// TIA Portal V17 export
// export: Created 2025-07-10T10:56:05.3982501Z, ExportSetting WithDefaults, DisplayName Totally Integrated Automation Portal, DisplayVersion V17, DisplayName TIA Portal Openness, DisplayVersion V17, DisplayName TIA Portal Version Control Interface, DisplayVersion V17, DisplayName SINAMICS Startdrive Advanced, DisplayVersion V17, DisplayName SINAMICS Startdrive G130, G150, S120, S150, SINAMICS MV, S210, DisplayVersion V17, DisplayName SINAMICS Startdrive G110M, G120, G120C, G120D, G120P, G115D, DisplayVersion V17, DisplayName STEP 7 Professional, DisplayVersion V17, DisplayName STEP 7 Safety, DisplayVersion V17, DisplayName WinCC Professional, DisplayVersion V17
FUNCTION_BLOCK "PR_GantryUnload_Seqv2 5_d22cba"   // FB1, LAD
VERSION : 0.1
// stored: AutoNumber true, IsIECCheckEnabled false, UDAEnableTagReadback false
   VAR_INPUT
      iAutoRunning : Bool;
      iCenteringSlideAtHome : Bool;
      iDistSenHighLimit : Int;
      iDistSenLowLimit : Int;
      iDistSensorIP : Int;
      iDryCycleWithoutPal : Bool;
      iGantryOutofZone : Bool;
      iGantryPickOver : Bool;
      iPCAckZero : Bool;
      iPCBypass : Bool;
      iPCDataReadOver : Bool;
      iPCDataWriteOver : Bool;
      iPalletPresent : Bool;
      iProcessStart : Bool;
      iReset_fault : Bool;
      iRetryPB : Bool;
      iScanErr : Bool;
      iScanOver : Bool;
      iScannerBypass : Bool;
      iSstMode : Bool;
      iSstPB : Bool;
   END_VAR
   VAR_OUTPUT
      qCenteringSlideAdvance : Bool;
      qCenteringSlideRetract : Bool;
      qCheckDistance : Bool;
      qGantryOkToUnload : Bool;
      qMsg : Array[0..2] of Bool;
      qPCReadCmd : Bool;
      qPCUploadCmd : Bool;
      qProcessOver : Bool;
      qScanCmd : Bool;
   END_VAR
   VAR DB_SPECIFIC
      StateNo : Int;
      s44_WaitResetRelease : Bool;
      s44_WaitResetRelease_T1 : Bool;
      s45_WaitGantryOutZone : Bool;
      s45_WaitGantryOutZone_T1 : Bool;
      s46_ChkStationHome : Bool;
      s46_ChkStationHome_T1 : Bool;
      s46_ChkStationHome_T2 : Bool;
      s47_WaitProcStartPZR : Bool;
      s47_WaitProcStartPZR_T1 : Bool;
      s48_ChkRecovery : Bool;
      s48_ChkRecovery_T1 : Bool;
      s48_ChkRecovery_T2 : Bool;
      s48_ChkRecovery_T3 : Bool;
      s49_WaitCentSlideAdv : Bool;
      s49_WaitCentSlideAdv_T1 : Bool;
      s50_WaitDistSensorFB : Bool;
      s50_WaitDistSensorFB_T1 : Bool;
      s51_WaitCentSlideRet : Bool;
      s51_WaitCentSlideRet_T1 : Bool;
      s52_WaitScanOver : Bool;
      s52_WaitScanOver_T1 : Bool;
      s52_WaitScanOver_T2 : Bool;
      s53_ChkMeasDistPCDat : Bool;
      s53_ChkMeasDistPCDat_T1 : Bool;
      s53_ChkMeasDistPCDat_T2 : Bool;
      s54_WaitGantryUnload : Bool;
      s54_WaitGantryUnload_T1 : Bool;
      s55_WaitGantryUnldOvr : Bool;
      s55_WaitGantryUnldOvr_T1 : Bool;
      s56_WaitGantryOutZone : Bool;
      s56_WaitGantryOutZone_T1 : Bool;
      s57_ChkReelAbsentCnv : Bool;
      s57_ChkReelAbsentCnv_T1 : Bool;
      s58_WaitProcStartLow : Bool;
      s58_WaitProcStartLow_T1 : Bool;
      s61_ChkMeasDiamTol : Bool;
      s61_ChkMeasDiamTol_T1 : Bool;
      s61_ChkMeasDiamTol_T2 : Bool;
      s62_WaitPCAckZero : Bool;
      s62_WaitPCAckZero_T1 : Bool;
      s63_WaitDataWritePC : Bool;
      s63_WaitDataWritePC_T1 : Bool;
      s64_WaitOperatorIntv : Bool;
      s64_WaitOperatorIntv_T1 : Bool;
      s65_ChkScanRetryOver : Bool;
      s65_ChkScanRetryOver_T1 : Bool;
      s65_ChkScanRetryOver_T2 : Bool;
      s66_WaitOperatorDecn : Bool;
      s66_WaitOperatorDecn_T1 : Bool;
      s67_WaitCentSlideRet : Bool;
      s67_WaitCentSlideRet_T1 : Bool;
      s68_WaitPCAckZeroRd : Bool;
      s68_WaitPCAckZeroRd_T1 : Bool;
      s69_WaitDataReadPC : Bool;
      s69_WaitDataReadPC_T1 : Bool;
      sDistanceHighLimit : Int;
      sDistanceLowLimit : Int;
      sRecoveryInt : Int;
      sScanRetryCount : Int;
      sSst : Bool;
      sSstPulse : Bool;
      sSstRise : Bool;
   END_VAR
   VAR_TEMP
      tOne : Bool;
   END_VAR
   VAR_TEMP   // added for the SCL form of the ladder/FBD networks
      _w1 : Bool;
   END_VAR
BEGIN

REGION Network 1
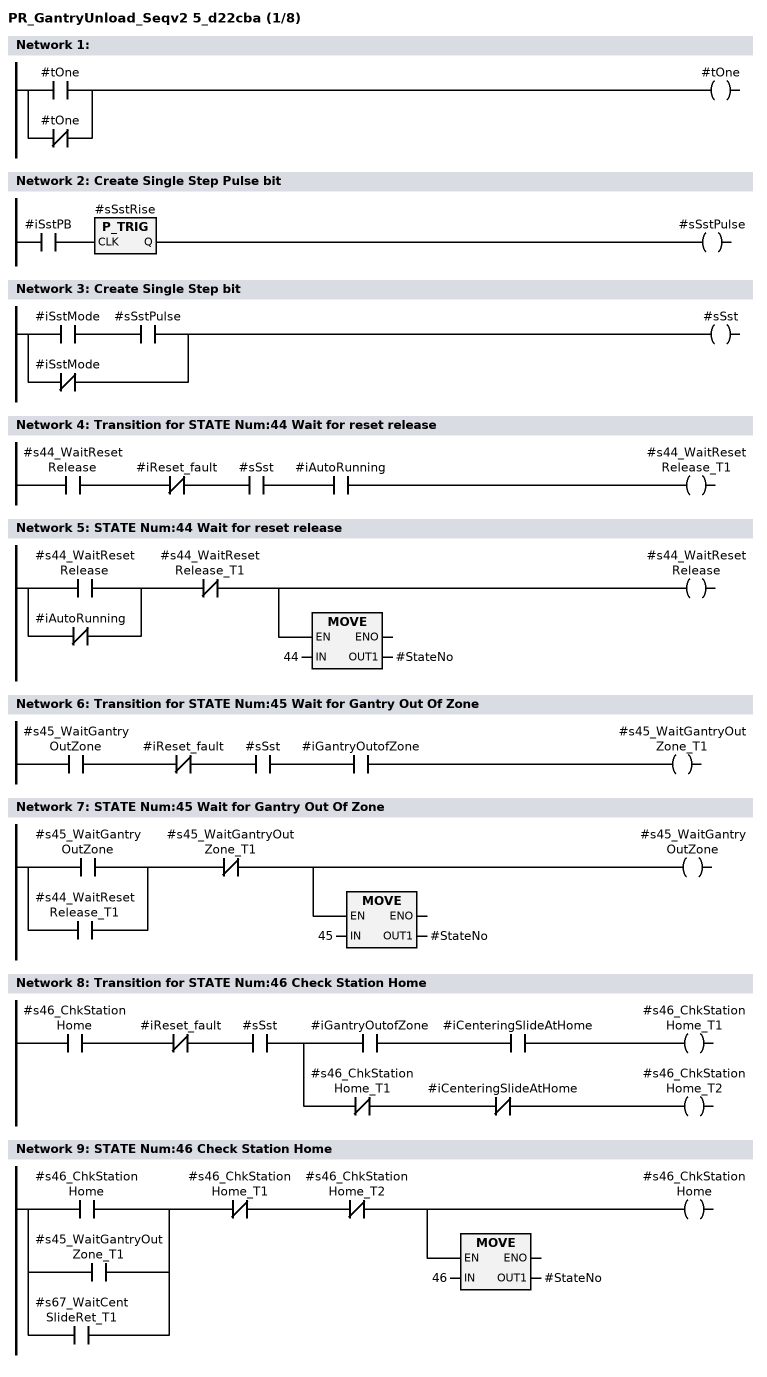
   RUNG wire#powerrail
      Contact( #tOne )
      wire#w1
      Coil( #tOne )
   END_RUNG
   RUNG wire#powerrail
      I_Contact( #tOne )
   END_RUNG wire#w1
   // the same network as SCL:
   #tOne := #tOne OR NOT #tOne;
END_REGION

REGION Network 2: Create Single Step Pulse bit
   RUNG wire#powerrail
      Contact( #iSstPB )
      P_Trig( #sSstRise )
      Coil( #sSstPulse )
   END_RUNG
   // the same network as SCL:
   #_w1 := #iSstPB AND NOT #sSstRise;   // rising edge
   #sSstRise := #iSstPB;
   #sSstPulse := #_w1;
END_REGION

REGION Network 3: Create Single Step bit
   RUNG wire#powerrail
      Contact( #iSstMode )
      Contact( #sSstPulse )
      wire#w1
      Coil( #sSst )
   END_RUNG
   RUNG wire#powerrail
      I_Contact( #iSstMode )
   END_RUNG wire#w1
   // the same network as SCL:
   #sSst := (#iSstMode AND #sSstPulse) OR NOT #iSstMode;
END_REGION

REGION Network 4: Transition for STATE Num:44 Wait for reset release
   RUNG wire#powerrail
      Contact( #s44_WaitResetRelease )
      I_Contact( #iReset_fault )
      Contact( #sSst )
      Contact( #iAutoRunning )
      Coil( #s44_WaitResetRelease_T1 )
   END_RUNG
   // the same network as SCL:
   #s44_WaitResetRelease_T1 := #s44_WaitResetRelease AND NOT #iReset_fault AND #sSst AND #iAutoRunning;
END_REGION

REGION Network 5: STATE Num:44 Wait for reset release
   RUNG wire#powerrail
      Contact( #s44_WaitResetRelease )
      wire#w1
      I_Contact( #s44_WaitResetRelease_T1 )
      wire#w2
      Coil( #s44_WaitResetRelease )
   END_RUNG
   RUNG wire#powerrail
      I_Contact( #iAutoRunning )
   END_RUNG wire#w1
   RUNG wire#w2
      { S7_GenerateENO := "TRUE" } Move(in := 44, out1 => #StateNo)
   END_RUNG
   // the same network as SCL:
   #s44_WaitResetRelease := (#s44_WaitResetRelease OR NOT #iAutoRunning) AND NOT #s44_WaitResetRelease_T1;
   IF #s44_WaitResetRelease THEN #StateNo := 44; END_IF;
END_REGION

REGION Network 6: Transition for STATE Num:45 Wait for Gantry Out Of Zone
   RUNG wire#powerrail
      Contact( #s45_WaitGantryOutZone )
      I_Contact( #iReset_fault )
      Contact( #sSst )
      Contact( #iGantryOutofZone )
      Coil( #s45_WaitGantryOutZone_T1 )
   END_RUNG
   // the same network as SCL:
   #s45_WaitGantryOutZone_T1 := #s45_WaitGantryOutZone AND NOT #iReset_fault AND #sSst AND #iGantryOutofZone;
END_REGION

REGION Network 7: STATE Num:45 Wait for Gantry Out Of Zone
   RUNG wire#powerrail
      Contact( #s45_WaitGantryOutZone )
      wire#w1
      I_Contact( #s45_WaitGantryOutZone_T1 )
      wire#w2
      Coil( #s45_WaitGantryOutZone )
   END_RUNG
   RUNG wire#powerrail
      Contact( #s44_WaitResetRelease_T1 )
   END_RUNG wire#w1
   RUNG wire#w2
      { S7_GenerateENO := "TRUE" } Move(in := 45, out1 => #StateNo)
   END_RUNG
   // the same network as SCL:
   #s45_WaitGantryOutZone := (#s45_WaitGantryOutZone OR #s44_WaitResetRelease_T1) AND NOT #s45_WaitGantryOutZone_T1;
   IF #s45_WaitGantryOutZone THEN #StateNo := 45; END_IF;
END_REGION

REGION Network 8: Transition for STATE Num:46 Check Station Home
   RUNG wire#powerrail
      Contact( #s46_ChkStationHome )
      I_Contact( #iReset_fault )
      Contact( #sSst )
      wire#w1
      Contact( #iGantryOutofZone )
      Contact( #iCenteringSlideAtHome )
      Coil( #s46_ChkStationHome_T1 )
   END_RUNG
   RUNG wire#w1
      I_Contact( #s46_ChkStationHome_T1 )
      I_Contact( #iCenteringSlideAtHome )
      Coil( #s46_ChkStationHome_T2 )
   END_RUNG
   // the same network as SCL:
   #_w1 := #s46_ChkStationHome AND NOT #iReset_fault AND #sSst;
   #s46_ChkStationHome_T1 := #_w1 AND #iGantryOutofZone AND #iCenteringSlideAtHome;
   #s46_ChkStationHome_T2 := #_w1 AND NOT #s46_ChkStationHome_T1 AND NOT #iCenteringSlideAtHome;
END_REGION

REGION Network 9: STATE Num:46 Check Station Home
   RUNG wire#powerrail
      Contact( #s46_ChkStationHome )
      wire#w1
      I_Contact( #s46_ChkStationHome_T1 )
      I_Contact( #s46_ChkStationHome_T2 )
      wire#w2
      Coil( #s46_ChkStationHome )
   END_RUNG
   RUNG wire#powerrail
      Contact( #s45_WaitGantryOutZone_T1 )
   END_RUNG wire#w1
   RUNG wire#powerrail
      Contact( #s67_WaitCentSlideRet_T1 )
   END_RUNG wire#w1
   RUNG wire#w2
      { S7_GenerateENO := "TRUE" } Move(in := 46, out1 => #StateNo)
   END_RUNG
   // the same network as SCL:
   #s46_ChkStationHome := (#s46_ChkStationHome OR #s45_WaitGantryOutZone_T1 OR #s67_WaitCentSlideRet_T1) AND NOT #s46_ChkStationHome_T1 AND NOT #s46_ChkStationHome_T2;
   IF #s46_ChkStationHome THEN #StateNo := 46; END_IF;
END_REGION

REGION Network 10: Transition for STATE Num:47 Wait for Process Start From PZR
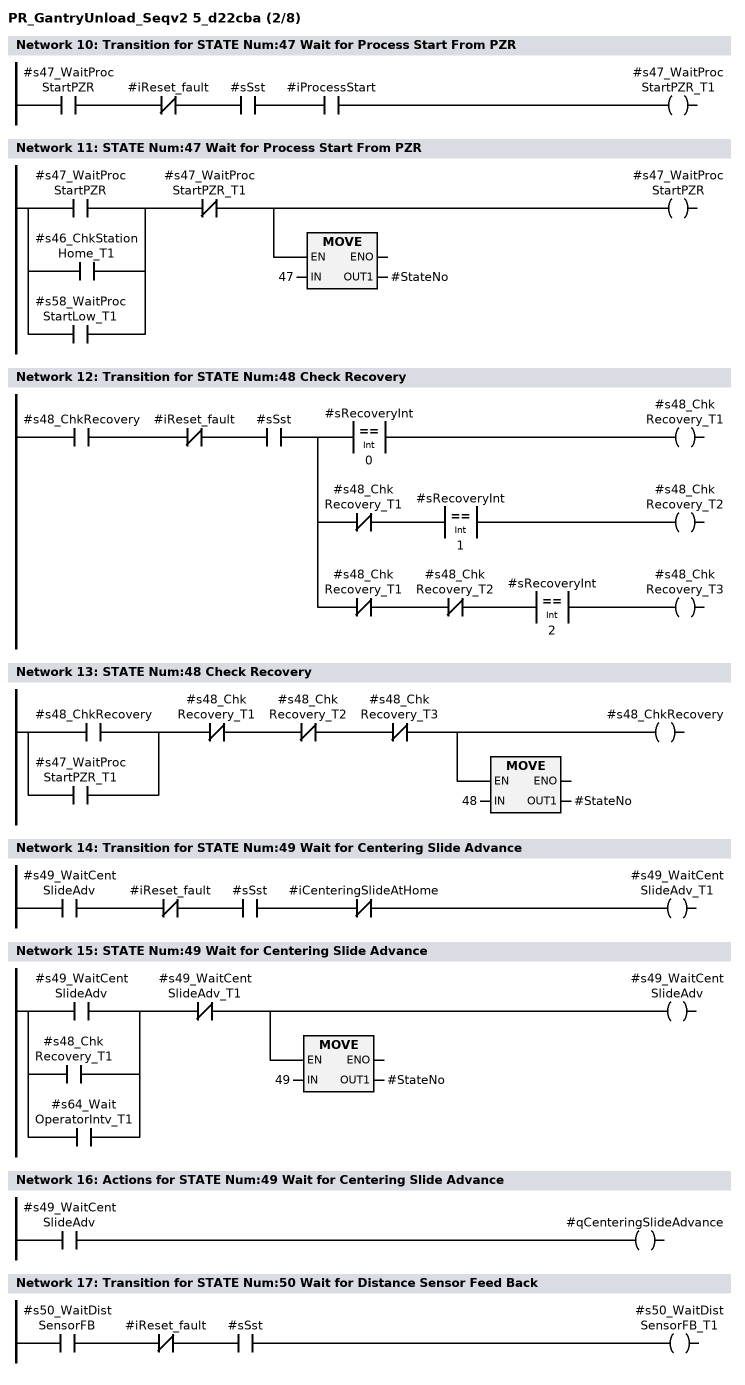
   RUNG wire#powerrail
      Contact( #s47_WaitProcStartPZR )
      I_Contact( #iReset_fault )
      Contact( #sSst )
      Contact( #iProcessStart )
      Coil( #s47_WaitProcStartPZR_T1 )
   END_RUNG
   // the same network as SCL:
   #s47_WaitProcStartPZR_T1 := #s47_WaitProcStartPZR AND NOT #iReset_fault AND #sSst AND #iProcessStart;
END_REGION

REGION Network 11: STATE Num:47 Wait for Process Start From PZR
   RUNG wire#powerrail
      Contact( #s47_WaitProcStartPZR )
      wire#w1
      I_Contact( #s47_WaitProcStartPZR_T1 )
      wire#w2
      Coil( #s47_WaitProcStartPZR )
   END_RUNG
   RUNG wire#powerrail
      Contact( #s46_ChkStationHome_T1 )
   END_RUNG wire#w1
   RUNG wire#powerrail
      Contact( #s58_WaitProcStartLow_T1 )
   END_RUNG wire#w1
   RUNG wire#w2
      { S7_GenerateENO := "TRUE" } Move(in := 47, out1 => #StateNo)
   END_RUNG
   // the same network as SCL:
   #s47_WaitProcStartPZR := (#s47_WaitProcStartPZR OR #s46_ChkStationHome_T1 OR #s58_WaitProcStartLow_T1) AND NOT #s47_WaitProcStartPZR_T1;
   IF #s47_WaitProcStartPZR THEN #StateNo := 47; END_IF;
END_REGION

REGION Network 12: Transition for STATE Num:48 Check Recovery
   RUNG wire#powerrail
      Contact( #s48_ChkRecovery )
      I_Contact( #iReset_fault )
      Contact( #sSst )
      wire#w1
      { S7_Templates := "SrcType := Int" } EQ_Contact(in1 := #sRecoveryInt, in2 := 0)
      Coil( #s48_ChkRecovery_T1 )
   END_RUNG
   RUNG wire#w1
      I_Contact( #s48_ChkRecovery_T1 )
      { S7_Templates := "SrcType := Int" } EQ_Contact(in1 := #sRecoveryInt, in2 := 1)
      Coil( #s48_ChkRecovery_T2 )
   END_RUNG
   RUNG wire#w1
      I_Contact( #s48_ChkRecovery_T1 )
      I_Contact( #s48_ChkRecovery_T2 )
      { S7_Templates := "SrcType := Int" } EQ_Contact(in1 := #sRecoveryInt, in2 := 2)
      Coil( #s48_ChkRecovery_T3 )
   END_RUNG
   // the same network as SCL:
   #_w1 := #s48_ChkRecovery AND NOT #iReset_fault AND #sSst;
   #s48_ChkRecovery_T1 := #_w1 AND (#sRecoveryInt = 0);
   #s48_ChkRecovery_T2 := #_w1 AND NOT #s48_ChkRecovery_T1 AND (#sRecoveryInt = 1);
   #s48_ChkRecovery_T3 := #_w1 AND NOT #s48_ChkRecovery_T1 AND NOT #s48_ChkRecovery_T2 AND (#sRecoveryInt = 2);
END_REGION

REGION Network 13: STATE Num:48 Check Recovery
   RUNG wire#powerrail
      Contact( #s48_ChkRecovery )
      wire#w1
      I_Contact( #s48_ChkRecovery_T1 )
      I_Contact( #s48_ChkRecovery_T2 )
      I_Contact( #s48_ChkRecovery_T3 )
      wire#w2
      Coil( #s48_ChkRecovery )
   END_RUNG
   RUNG wire#powerrail
      Contact( #s47_WaitProcStartPZR_T1 )
   END_RUNG wire#w1
   RUNG wire#w2
      { S7_GenerateENO := "TRUE" } Move(in := 48, out1 => #StateNo)
   END_RUNG
   // the same network as SCL:
   #s48_ChkRecovery := (#s48_ChkRecovery OR #s47_WaitProcStartPZR_T1) AND NOT #s48_ChkRecovery_T1 AND NOT #s48_ChkRecovery_T2 AND NOT #s48_ChkRecovery_T3;
   IF #s48_ChkRecovery THEN #StateNo := 48; END_IF;
END_REGION

REGION Network 14: Transition for STATE Num:49 Wait for Centering Slide Advance
   RUNG wire#powerrail
      Contact( #s49_WaitCentSlideAdv )
      I_Contact( #iReset_fault )
      Contact( #sSst )
      I_Contact( #iCenteringSlideAtHome )
      Coil( #s49_WaitCentSlideAdv_T1 )
   END_RUNG
   // the same network as SCL:
   #s49_WaitCentSlideAdv_T1 := #s49_WaitCentSlideAdv AND NOT #iReset_fault AND #sSst AND NOT #iCenteringSlideAtHome;
END_REGION

REGION Network 15: STATE Num:49 Wait for Centering Slide Advance
   RUNG wire#powerrail
      Contact( #s49_WaitCentSlideAdv )
      wire#w1
      I_Contact( #s49_WaitCentSlideAdv_T1 )
      wire#w2
      Coil( #s49_WaitCentSlideAdv )
   END_RUNG
   RUNG wire#powerrail
      Contact( #s48_ChkRecovery_T1 )
   END_RUNG wire#w1
   RUNG wire#powerrail
      Contact( #s64_WaitOperatorIntv_T1 )
   END_RUNG wire#w1
   RUNG wire#w2
      { S7_GenerateENO := "TRUE" } Move(in := 49, out1 => #StateNo)
   END_RUNG
   // the same network as SCL:
   #s49_WaitCentSlideAdv := (#s49_WaitCentSlideAdv OR #s48_ChkRecovery_T1 OR #s64_WaitOperatorIntv_T1) AND NOT #s49_WaitCentSlideAdv_T1;
   IF #s49_WaitCentSlideAdv THEN #StateNo := 49; END_IF;
END_REGION

REGION Network 16: Actions for STATE Num:49 Wait for Centering Slide Advance
   RUNG wire#powerrail
      Contact( #s49_WaitCentSlideAdv )
      Coil( #qCenteringSlideAdvance )
   END_RUNG
   // the same network as SCL:
   #qCenteringSlideAdvance := #s49_WaitCentSlideAdv;
END_REGION

REGION Network 17: Transition for STATE Num:50 Wait for Distance Sensor Feed Back
   RUNG wire#powerrail
      Contact( #s50_WaitDistSensorFB )
      I_Contact( #iReset_fault )
      Contact( #sSst )
      Coil( #s50_WaitDistSensorFB_T1 )
   END_RUNG
   // the same network as SCL:
   #s50_WaitDistSensorFB_T1 := #s50_WaitDistSensorFB AND NOT #iReset_fault AND #sSst;
END_REGION

REGION Network 18: STATE Num:50 Wait for Distance Sensor Feed Back
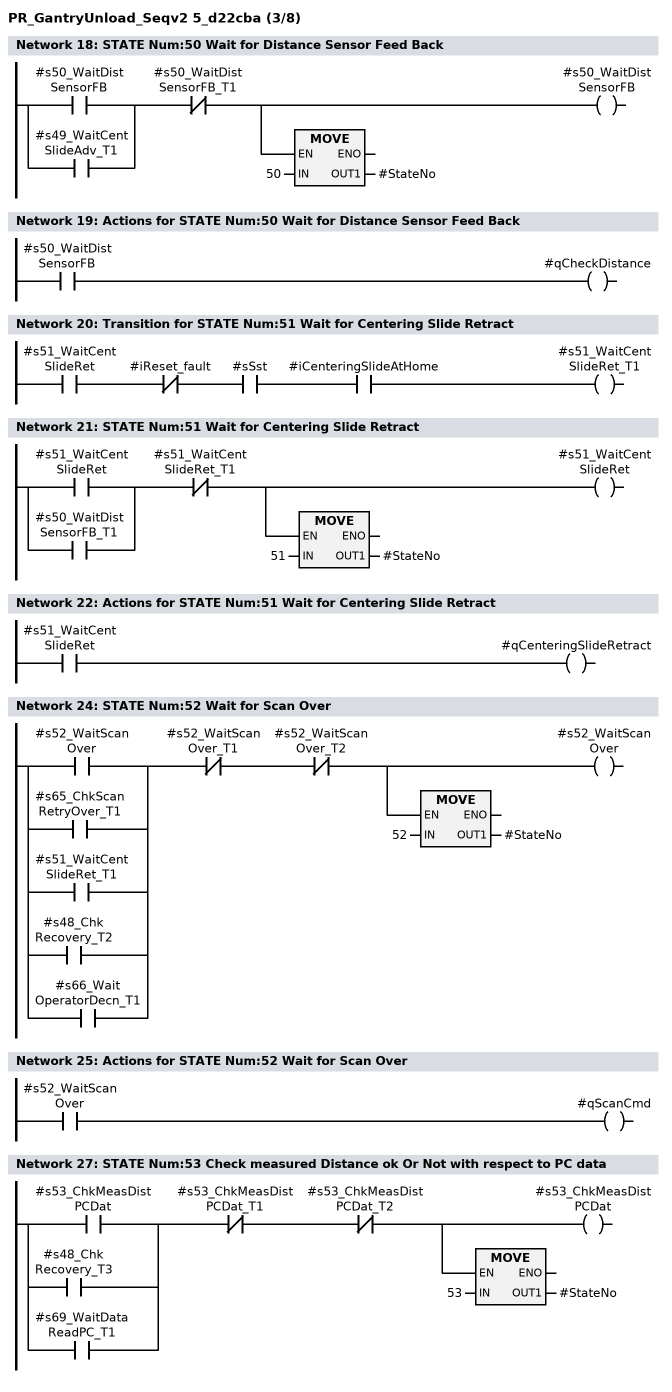
   RUNG wire#powerrail
      Contact( #s50_WaitDistSensorFB )
      wire#w1
      I_Contact( #s50_WaitDistSensorFB_T1 )
      wire#w2
      Coil( #s50_WaitDistSensorFB )
   END_RUNG
   RUNG wire#powerrail
      Contact( #s49_WaitCentSlideAdv_T1 )
   END_RUNG wire#w1
   RUNG wire#w2
      { S7_GenerateENO := "TRUE" } Move(in := 50, out1 => #StateNo)
   END_RUNG
   // the same network as SCL:
   #s50_WaitDistSensorFB := (#s50_WaitDistSensorFB OR #s49_WaitCentSlideAdv_T1) AND NOT #s50_WaitDistSensorFB_T1;
   IF #s50_WaitDistSensorFB THEN #StateNo := 50; END_IF;
END_REGION

REGION Network 19: Actions for STATE Num:50 Wait for Distance Sensor Feed Back
   RUNG wire#powerrail
      Contact( #s50_WaitDistSensorFB )
      Coil( #qCheckDistance )
   END_RUNG
   // the same network as SCL:
   #qCheckDistance := #s50_WaitDistSensorFB;
END_REGION

REGION Network 20: Transition for STATE Num:51 Wait for Centering Slide Retract
   RUNG wire#powerrail
      Contact( #s51_WaitCentSlideRet )
      I_Contact( #iReset_fault )
      Contact( #sSst )
      Contact( #iCenteringSlideAtHome )
      Coil( #s51_WaitCentSlideRet_T1 )
   END_RUNG
   // the same network as SCL:
   #s51_WaitCentSlideRet_T1 := #s51_WaitCentSlideRet AND NOT #iReset_fault AND #sSst AND #iCenteringSlideAtHome;
END_REGION

REGION Network 21: STATE Num:51 Wait for Centering Slide Retract
   RUNG wire#powerrail
      Contact( #s51_WaitCentSlideRet )
      wire#w1
      I_Contact( #s51_WaitCentSlideRet_T1 )
      wire#w2
      Coil( #s51_WaitCentSlideRet )
   END_RUNG
   RUNG wire#powerrail
      Contact( #s50_WaitDistSensorFB_T1 )
   END_RUNG wire#w1
   RUNG wire#w2
      { S7_GenerateENO := "TRUE" } Move(in := 51, out1 => #StateNo)
   END_RUNG
   // the same network as SCL:
   #s51_WaitCentSlideRet := (#s51_WaitCentSlideRet OR #s50_WaitDistSensorFB_T1) AND NOT #s51_WaitCentSlideRet_T1;
   IF #s51_WaitCentSlideRet THEN #StateNo := 51; END_IF;
END_REGION

REGION Network 22: Actions for STATE Num:51 Wait for Centering Slide Retract
   RUNG wire#powerrail
      Contact( #s51_WaitCentSlideRet )
      Coil( #qCenteringSlideRetract )
   END_RUNG
   // the same network as SCL:
   #qCenteringSlideRetract := #s51_WaitCentSlideRet;
END_REGION

NETWORK
TITLE = Transition for STATE Num:52 Wait for Scan Over
      A     #s52_WaitScanOver;
      AN    #iReset_fault;
      A     #sSst;
      =     %L1.0;
      A     %L1.0;
      A(;
      O     #iScanOver;
      AN    #iScanErr;
      );
      O     #iScannerBypass;
      O     #iDryCycleWithoutPal;
      =     #s52_WaitScanOver_T1;
      A     %L1.0;
      AN    #s52_WaitScanOver_T1;
      A     #iScanErr;
      =     #s52_WaitScanOver_T2;

REGION Network 24: STATE Num:52 Wait for Scan Over
   RUNG wire#powerrail
      Contact( #s52_WaitScanOver )
      wire#w1
      I_Contact( #s52_WaitScanOver_T1 )
      I_Contact( #s52_WaitScanOver_T2 )
      wire#w2
      Coil( #s52_WaitScanOver )
   END_RUNG
   RUNG wire#powerrail
      Contact( #s65_ChkScanRetryOver_T1 )
   END_RUNG wire#w1
   RUNG wire#powerrail
      Contact( #s51_WaitCentSlideRet_T1 )
   END_RUNG wire#w1
   RUNG wire#powerrail
      Contact( #s48_ChkRecovery_T2 )
   END_RUNG wire#w1
   RUNG wire#powerrail
      Contact( #s66_WaitOperatorDecn_T1 )
   END_RUNG wire#w1
   RUNG wire#w2
      { S7_GenerateENO := "TRUE" } Move(in := 52, out1 => #StateNo)
   END_RUNG
   // the same network as SCL:
   #s52_WaitScanOver := (#s52_WaitScanOver OR #s65_ChkScanRetryOver_T1 OR #s51_WaitCentSlideRet_T1 OR #s48_ChkRecovery_T2 OR #s66_WaitOperatorDecn_T1) AND NOT #s52_WaitScanOver_T1 AND NOT #s52_WaitScanOver_T2;
   IF #s52_WaitScanOver THEN #StateNo := 52; END_IF;
END_REGION

REGION Network 25: Actions for STATE Num:52 Wait for Scan Over
   RUNG wire#powerrail
      Contact( #s52_WaitScanOver )
      Coil( #qScanCmd )
   END_RUNG
   // the same network as SCL:
   #qScanCmd := #s52_WaitScanOver;
END_REGION

NETWORK
TITLE = Transition for STATE Num:53 Check measured Distance ok Or Not with respect to PC data
      A     #s53_ChkMeasDistPCDat;
      AN    #iReset_fault;
      A     #sSst;
      =     %L1.0;
      A     %L1.0;
      A(;
      L     #iDistSensorIP;
      L     #sDistanceLowLimit;
      >=R;
      );
      O(;
      L     #iDistSensorIP;
      L     #sDistanceHighLimit;
      <=R;
      );
      =     #s53_ChkMeasDistPCDat_T1;
      A     %L1.0;
      AN    #s53_ChkMeasDistPCDat_T1;
      A(;
      L     #iDistSensorIP;
      L     #sDistanceLowLimit;
      <R;
      );
      O(;
      L     #iDistSensorIP;
      L     #sDistanceHighLimit;
      >R;
      );
      =     #s53_ChkMeasDistPCDat_T2;

REGION Network 27: STATE Num:53 Check measured Distance ok Or Not with respect to PC data
   RUNG wire#powerrail
      Contact( #s53_ChkMeasDistPCDat )
      wire#w1
      I_Contact( #s53_ChkMeasDistPCDat_T1 )
      I_Contact( #s53_ChkMeasDistPCDat_T2 )
      wire#w2
      Coil( #s53_ChkMeasDistPCDat )
   END_RUNG
   RUNG wire#powerrail
      Contact( #s48_ChkRecovery_T3 )
   END_RUNG wire#w1
   RUNG wire#powerrail
      Contact( #s69_WaitDataReadPC_T1 )
   END_RUNG wire#w1
   RUNG wire#w2
      { S7_GenerateENO := "TRUE" } Move(in := 53, out1 => #StateNo)
   END_RUNG
   // the same network as SCL:
   #s53_ChkMeasDistPCDat := (#s53_ChkMeasDistPCDat OR #s48_ChkRecovery_T3 OR #s69_WaitDataReadPC_T1) AND NOT #s53_ChkMeasDistPCDat_T1 AND NOT #s53_ChkMeasDistPCDat_T2;
   IF #s53_ChkMeasDistPCDat THEN #StateNo := 53; END_IF;
END_REGION

REGION Network 28: Transition for STATE Num:54 Wait for Gantry at Unload Position.
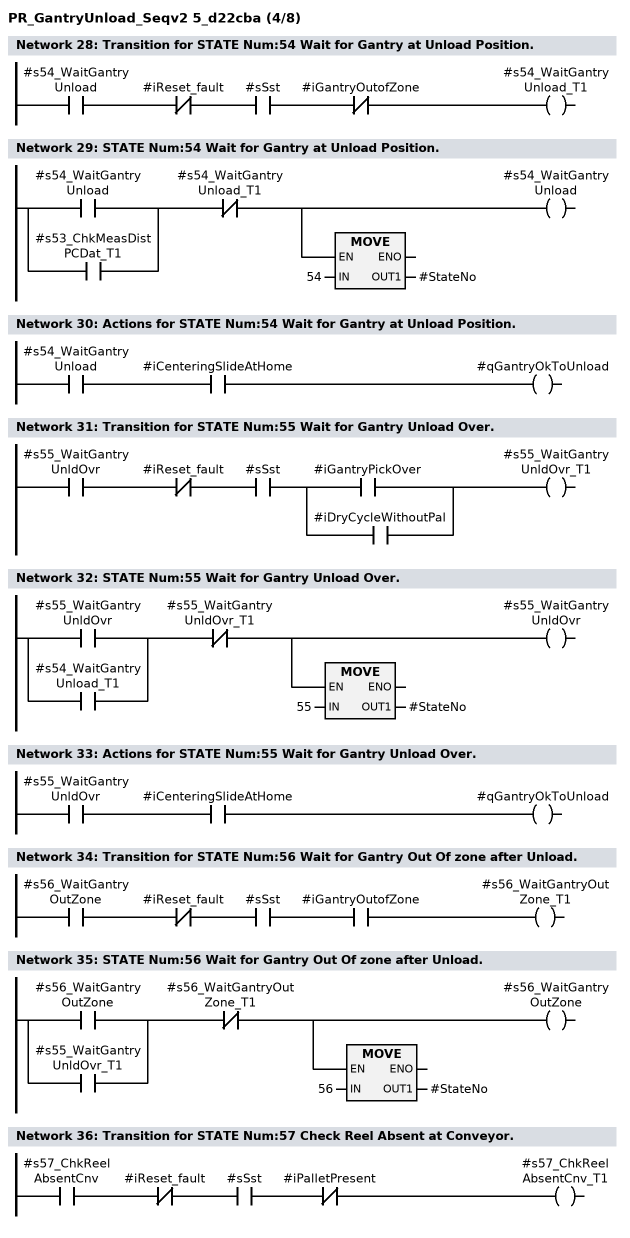
   RUNG wire#powerrail
      Contact( #s54_WaitGantryUnload )
      I_Contact( #iReset_fault )
      Contact( #sSst )
      I_Contact( #iGantryOutofZone )
      Coil( #s54_WaitGantryUnload_T1 )
   END_RUNG
   // the same network as SCL:
   #s54_WaitGantryUnload_T1 := #s54_WaitGantryUnload AND NOT #iReset_fault AND #sSst AND NOT #iGantryOutofZone;
END_REGION

REGION Network 29: STATE Num:54 Wait for Gantry at Unload Position.
   RUNG wire#powerrail
      Contact( #s54_WaitGantryUnload )
      wire#w1
      I_Contact( #s54_WaitGantryUnload_T1 )
      wire#w2
      Coil( #s54_WaitGantryUnload )
   END_RUNG
   RUNG wire#powerrail
      Contact( #s53_ChkMeasDistPCDat_T1 )
   END_RUNG wire#w1
   RUNG wire#w2
      { S7_GenerateENO := "TRUE" } Move(in := 54, out1 => #StateNo)
   END_RUNG
   // the same network as SCL:
   #s54_WaitGantryUnload := (#s54_WaitGantryUnload OR #s53_ChkMeasDistPCDat_T1) AND NOT #s54_WaitGantryUnload_T1;
   IF #s54_WaitGantryUnload THEN #StateNo := 54; END_IF;
END_REGION

REGION Network 30: Actions for STATE Num:54 Wait for Gantry at Unload Position.
   RUNG wire#powerrail
      Contact( #s54_WaitGantryUnload )
      Contact( #iCenteringSlideAtHome )
      Coil( #qGantryOkToUnload )
   END_RUNG
   // the same network as SCL:
   #qGantryOkToUnload := #s54_WaitGantryUnload AND #iCenteringSlideAtHome;
END_REGION

REGION Network 31: Transition for STATE Num:55 Wait for Gantry Unload Over.
   RUNG wire#powerrail
      Contact( #s55_WaitGantryUnldOvr )
      I_Contact( #iReset_fault )
      Contact( #sSst )
      wire#w1
      Contact( #iGantryPickOver )
      wire#w2
      Coil( #s55_WaitGantryUnldOvr_T1 )
   END_RUNG
   RUNG wire#w1
      Contact( #iDryCycleWithoutPal )
   END_RUNG wire#w2
   // the same network as SCL:
   #s55_WaitGantryUnldOvr_T1 := #s55_WaitGantryUnldOvr AND NOT #iReset_fault AND #sSst AND (#iGantryPickOver OR #iDryCycleWithoutPal);
END_REGION

REGION Network 32: STATE Num:55 Wait for Gantry Unload Over.
   RUNG wire#powerrail
      Contact( #s55_WaitGantryUnldOvr )
      wire#w1
      I_Contact( #s55_WaitGantryUnldOvr_T1 )
      wire#w2
      Coil( #s55_WaitGantryUnldOvr )
   END_RUNG
   RUNG wire#powerrail
      Contact( #s54_WaitGantryUnload_T1 )
   END_RUNG wire#w1
   RUNG wire#w2
      { S7_GenerateENO := "TRUE" } Move(in := 55, out1 => #StateNo)
   END_RUNG
   // the same network as SCL:
   #s55_WaitGantryUnldOvr := (#s55_WaitGantryUnldOvr OR #s54_WaitGantryUnload_T1) AND NOT #s55_WaitGantryUnldOvr_T1;
   IF #s55_WaitGantryUnldOvr THEN #StateNo := 55; END_IF;
END_REGION

REGION Network 33: Actions for STATE Num:55 Wait for Gantry Unload Over.
   RUNG wire#powerrail
      Contact( #s55_WaitGantryUnldOvr )
      Contact( #iCenteringSlideAtHome )
      Coil( #qGantryOkToUnload )
   END_RUNG
   // the same network as SCL:
   #qGantryOkToUnload := #s55_WaitGantryUnldOvr AND #iCenteringSlideAtHome;
END_REGION

REGION Network 34: Transition for STATE Num:56 Wait for Gantry Out Of zone after Unload.
   RUNG wire#powerrail
      Contact( #s56_WaitGantryOutZone )
      I_Contact( #iReset_fault )
      Contact( #sSst )
      Contact( #iGantryOutofZone )
      Coil( #s56_WaitGantryOutZone_T1 )
   END_RUNG
   // the same network as SCL:
   #s56_WaitGantryOutZone_T1 := #s56_WaitGantryOutZone AND NOT #iReset_fault AND #sSst AND #iGantryOutofZone;
END_REGION

REGION Network 35: STATE Num:56 Wait for Gantry Out Of zone after Unload.
   RUNG wire#powerrail
      Contact( #s56_WaitGantryOutZone )
      wire#w1
      I_Contact( #s56_WaitGantryOutZone_T1 )
      wire#w2
      Coil( #s56_WaitGantryOutZone )
   END_RUNG
   RUNG wire#powerrail
      Contact( #s55_WaitGantryUnldOvr_T1 )
   END_RUNG wire#w1
   RUNG wire#w2
      { S7_GenerateENO := "TRUE" } Move(in := 56, out1 => #StateNo)
   END_RUNG
   // the same network as SCL:
   #s56_WaitGantryOutZone := (#s56_WaitGantryOutZone OR #s55_WaitGantryUnldOvr_T1) AND NOT #s56_WaitGantryOutZone_T1;
   IF #s56_WaitGantryOutZone THEN #StateNo := 56; END_IF;
END_REGION

REGION Network 36: Transition for STATE Num:57 Check Reel Absent at Conveyor.
   RUNG wire#powerrail
      Contact( #s57_ChkReelAbsentCnv )
      I_Contact( #iReset_fault )
      Contact( #sSst )
      I_Contact( #iPalletPresent )
      Coil( #s57_ChkReelAbsentCnv_T1 )
   END_RUNG
   // the same network as SCL:
   #s57_ChkReelAbsentCnv_T1 := #s57_ChkReelAbsentCnv AND NOT #iReset_fault AND #sSst AND NOT #iPalletPresent;
END_REGION

REGION Network 37: STATE Num:57 Check Reel Absent at Conveyor.
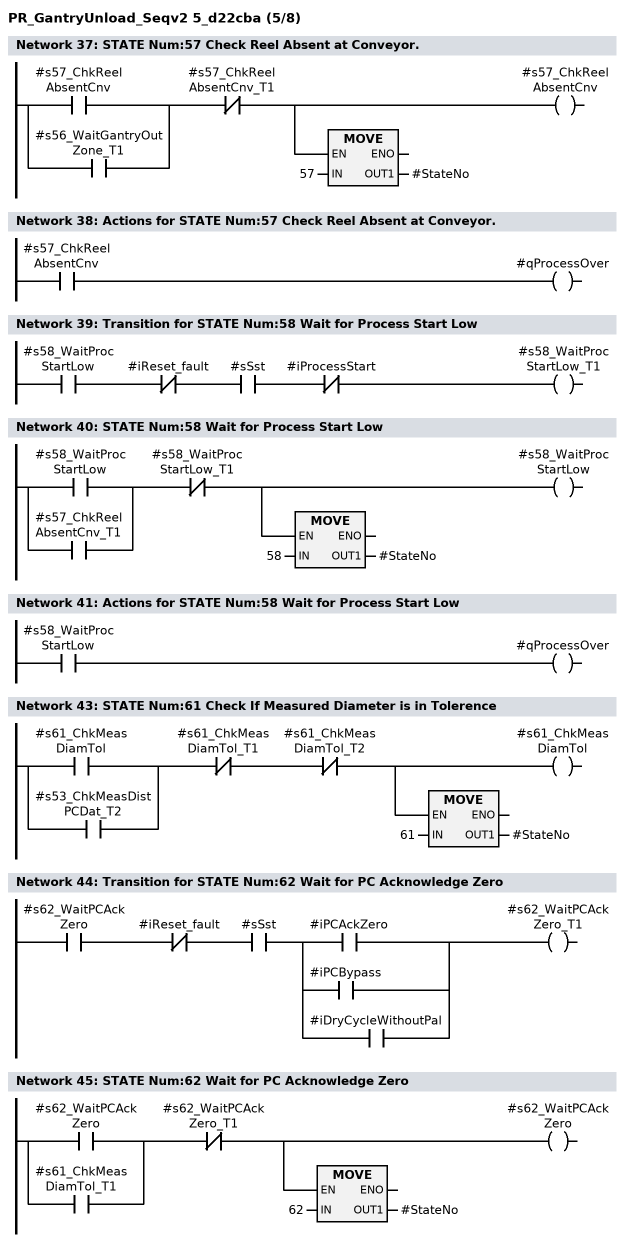
   RUNG wire#powerrail
      Contact( #s57_ChkReelAbsentCnv )
      wire#w1
      I_Contact( #s57_ChkReelAbsentCnv_T1 )
      wire#w2
      Coil( #s57_ChkReelAbsentCnv )
   END_RUNG
   RUNG wire#powerrail
      Contact( #s56_WaitGantryOutZone_T1 )
   END_RUNG wire#w1
   RUNG wire#w2
      { S7_GenerateENO := "TRUE" } Move(in := 57, out1 => #StateNo)
   END_RUNG
   // the same network as SCL:
   #s57_ChkReelAbsentCnv := (#s57_ChkReelAbsentCnv OR #s56_WaitGantryOutZone_T1) AND NOT #s57_ChkReelAbsentCnv_T1;
   IF #s57_ChkReelAbsentCnv THEN #StateNo := 57; END_IF;
END_REGION

REGION Network 38: Actions for STATE Num:57 Check Reel Absent at Conveyor.
   RUNG wire#powerrail
      Contact( #s57_ChkReelAbsentCnv )
      Coil( #qProcessOver )
   END_RUNG
   // the same network as SCL:
   #qProcessOver := #s57_ChkReelAbsentCnv;
END_REGION

REGION Network 39: Transition for STATE Num:58 Wait for Process Start Low
   RUNG wire#powerrail
      Contact( #s58_WaitProcStartLow )
      I_Contact( #iReset_fault )
      Contact( #sSst )
      I_Contact( #iProcessStart )
      Coil( #s58_WaitProcStartLow_T1 )
   END_RUNG
   // the same network as SCL:
   #s58_WaitProcStartLow_T1 := #s58_WaitProcStartLow AND NOT #iReset_fault AND #sSst AND NOT #iProcessStart;
END_REGION

REGION Network 40: STATE Num:58 Wait for Process Start Low
   RUNG wire#powerrail
      Contact( #s58_WaitProcStartLow )
      wire#w1
      I_Contact( #s58_WaitProcStartLow_T1 )
      wire#w2
      Coil( #s58_WaitProcStartLow )
   END_RUNG
   RUNG wire#powerrail
      Contact( #s57_ChkReelAbsentCnv_T1 )
   END_RUNG wire#w1
   RUNG wire#w2
      { S7_GenerateENO := "TRUE" } Move(in := 58, out1 => #StateNo)
   END_RUNG
   // the same network as SCL:
   #s58_WaitProcStartLow := (#s58_WaitProcStartLow OR #s57_ChkReelAbsentCnv_T1) AND NOT #s58_WaitProcStartLow_T1;
   IF #s58_WaitProcStartLow THEN #StateNo := 58; END_IF;
END_REGION

REGION Network 41: Actions for STATE Num:58 Wait for Process Start Low
   RUNG wire#powerrail
      Contact( #s58_WaitProcStartLow )
      Coil( #qProcessOver )
   END_RUNG
   // the same network as SCL:
   #qProcessOver := #s58_WaitProcStartLow;
END_REGION

NETWORK
TITLE = Transition for STATE Num:61 Check If Measured Diameter is in Tolerence
      A     #s61_ChkMeasDiamTol;
      AN    #iReset_fault;
      A     #sSst;
      =     %L1.0;
      A     %L1.0;
      A(;
      L     #iDistSenLowLimit;
      L     #iDistSensorIP;
      <=R;
      );
      O(;
      L     #iDistSensorIP;
      L     #iDistSenHighLimit;
      <=R;
      );
      =     #s61_ChkMeasDiamTol_T1;
      A     %L1.0;
      AN    #s61_ChkMeasDiamTol_T1;
      A(;
      L     #iDistSenLowLimit;
      L     #iDistSensorIP;
      >R;
      );
      O(;
      L     #iDistSensorIP;
      L     #iDistSenHighLimit;
      >R;
      );
      =     #s61_ChkMeasDiamTol_T2;

REGION Network 43: STATE Num:61 Check If Measured Diameter is in Tolerence
   RUNG wire#powerrail
      Contact( #s61_ChkMeasDiamTol )
      wire#w1
      I_Contact( #s61_ChkMeasDiamTol_T1 )
      I_Contact( #s61_ChkMeasDiamTol_T2 )
      wire#w2
      Coil( #s61_ChkMeasDiamTol )
   END_RUNG
   RUNG wire#powerrail
      Contact( #s53_ChkMeasDistPCDat_T2 )
   END_RUNG wire#w1
   RUNG wire#w2
      { S7_GenerateENO := "TRUE" } Move(in := 61, out1 => #StateNo)
   END_RUNG
   // the same network as SCL:
   #s61_ChkMeasDiamTol := (#s61_ChkMeasDiamTol OR #s53_ChkMeasDistPCDat_T2) AND NOT #s61_ChkMeasDiamTol_T1 AND NOT #s61_ChkMeasDiamTol_T2;
   IF #s61_ChkMeasDiamTol THEN #StateNo := 61; END_IF;
END_REGION

REGION Network 44: Transition for STATE Num:62 Wait for PC Acknowledge Zero
   RUNG wire#powerrail
      Contact( #s62_WaitPCAckZero )
      I_Contact( #iReset_fault )
      Contact( #sSst )
      wire#w1
      Contact( #iPCAckZero )
      wire#w2
      Coil( #s62_WaitPCAckZero_T1 )
   END_RUNG
   RUNG wire#w1
      Contact( #iPCBypass )
   END_RUNG wire#w2
   RUNG wire#w1
      Contact( #iDryCycleWithoutPal )
   END_RUNG wire#w2
   // the same network as SCL:
   #s62_WaitPCAckZero_T1 := #s62_WaitPCAckZero AND NOT #iReset_fault AND #sSst AND (#iPCAckZero OR #iPCBypass OR #iDryCycleWithoutPal);
END_REGION

REGION Network 45: STATE Num:62 Wait for PC Acknowledge Zero
   RUNG wire#powerrail
      Contact( #s62_WaitPCAckZero )
      wire#w1
      I_Contact( #s62_WaitPCAckZero_T1 )
      wire#w2
      Coil( #s62_WaitPCAckZero )
   END_RUNG
   RUNG wire#powerrail
      Contact( #s61_ChkMeasDiamTol_T1 )
   END_RUNG wire#w1
   RUNG wire#w2
      { S7_GenerateENO := "TRUE" } Move(in := 62, out1 => #StateNo)
   END_RUNG
   // the same network as SCL:
   #s62_WaitPCAckZero := (#s62_WaitPCAckZero OR #s61_ChkMeasDiamTol_T1) AND NOT #s62_WaitPCAckZero_T1;
   IF #s62_WaitPCAckZero THEN #StateNo := 62; END_IF;
END_REGION

REGION Network 46: Transition for STATE Num:63 Wait for Data Write Over From PC
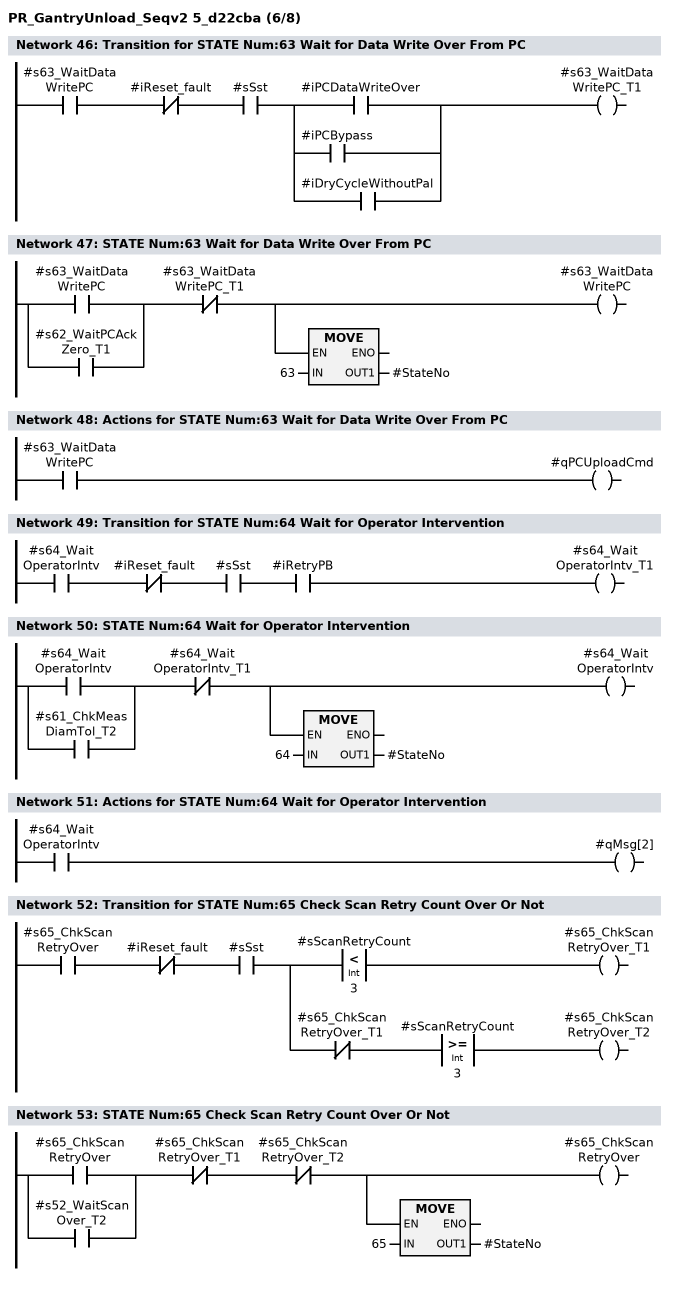
   RUNG wire#powerrail
      Contact( #s63_WaitDataWritePC )
      I_Contact( #iReset_fault )
      Contact( #sSst )
      wire#w1
      Contact( #iPCDataWriteOver )
      wire#w2
      Coil( #s63_WaitDataWritePC_T1 )
   END_RUNG
   RUNG wire#w1
      Contact( #iPCBypass )
   END_RUNG wire#w2
   RUNG wire#w1
      Contact( #iDryCycleWithoutPal )
   END_RUNG wire#w2
   // the same network as SCL:
   #s63_WaitDataWritePC_T1 := #s63_WaitDataWritePC AND NOT #iReset_fault AND #sSst AND (#iPCDataWriteOver OR #iPCBypass OR #iDryCycleWithoutPal);
END_REGION

REGION Network 47: STATE Num:63 Wait for Data Write Over From PC
   RUNG wire#powerrail
      Contact( #s63_WaitDataWritePC )
      wire#w1
      I_Contact( #s63_WaitDataWritePC_T1 )
      wire#w2
      Coil( #s63_WaitDataWritePC )
   END_RUNG
   RUNG wire#powerrail
      Contact( #s62_WaitPCAckZero_T1 )
   END_RUNG wire#w1
   RUNG wire#w2
      { S7_GenerateENO := "TRUE" } Move(in := 63, out1 => #StateNo)
   END_RUNG
   // the same network as SCL:
   #s63_WaitDataWritePC := (#s63_WaitDataWritePC OR #s62_WaitPCAckZero_T1) AND NOT #s63_WaitDataWritePC_T1;
   IF #s63_WaitDataWritePC THEN #StateNo := 63; END_IF;
END_REGION

REGION Network 48: Actions for STATE Num:63 Wait for Data Write Over From PC
   RUNG wire#powerrail
      Contact( #s63_WaitDataWritePC )
      Coil( #qPCUploadCmd )
   END_RUNG
   // the same network as SCL:
   #qPCUploadCmd := #s63_WaitDataWritePC;
END_REGION

REGION Network 49: Transition for STATE Num:64 Wait for Operator Intervention
   RUNG wire#powerrail
      Contact( #s64_WaitOperatorIntv )
      I_Contact( #iReset_fault )
      Contact( #sSst )
      Contact( #iRetryPB )
      Coil( #s64_WaitOperatorIntv_T1 )
   END_RUNG
   // the same network as SCL:
   #s64_WaitOperatorIntv_T1 := #s64_WaitOperatorIntv AND NOT #iReset_fault AND #sSst AND #iRetryPB;
END_REGION

REGION Network 50: STATE Num:64 Wait for Operator Intervention
   RUNG wire#powerrail
      Contact( #s64_WaitOperatorIntv )
      wire#w1
      I_Contact( #s64_WaitOperatorIntv_T1 )
      wire#w2
      Coil( #s64_WaitOperatorIntv )
   END_RUNG
   RUNG wire#powerrail
      Contact( #s61_ChkMeasDiamTol_T2 )
   END_RUNG wire#w1
   RUNG wire#w2
      { S7_GenerateENO := "TRUE" } Move(in := 64, out1 => #StateNo)
   END_RUNG
   // the same network as SCL:
   #s64_WaitOperatorIntv := (#s64_WaitOperatorIntv OR #s61_ChkMeasDiamTol_T2) AND NOT #s64_WaitOperatorIntv_T1;
   IF #s64_WaitOperatorIntv THEN #StateNo := 64; END_IF;
END_REGION

REGION Network 51: Actions for STATE Num:64 Wait for Operator Intervention
   RUNG wire#powerrail
      Contact( #s64_WaitOperatorIntv )
      Coil( #qMsg[2] )
   END_RUNG
   // the same network as SCL:
   #qMsg[2] := #s64_WaitOperatorIntv;
END_REGION

REGION Network 52: Transition for STATE Num:65 Check Scan Retry Count Over Or Not
   RUNG wire#powerrail
      Contact( #s65_ChkScanRetryOver )
      I_Contact( #iReset_fault )
      Contact( #sSst )
      wire#w1
      { S7_Templates := "SrcType := Int" } LT_Contact(in1 := #sScanRetryCount, in2 := 3)
      Coil( #s65_ChkScanRetryOver_T1 )
   END_RUNG
   RUNG wire#w1
      I_Contact( #s65_ChkScanRetryOver_T1 )
      { S7_Templates := "SrcType := Int" } GE_Contact(in1 := #sScanRetryCount, in2 := 3)
      Coil( #s65_ChkScanRetryOver_T2 )
   END_RUNG
   // the same network as SCL:
   #_w1 := #s65_ChkScanRetryOver AND NOT #iReset_fault AND #sSst;
   #s65_ChkScanRetryOver_T1 := #_w1 AND (#sScanRetryCount < 3);
   #s65_ChkScanRetryOver_T2 := #_w1 AND NOT #s65_ChkScanRetryOver_T1 AND (#sScanRetryCount >= 3);
END_REGION

REGION Network 53: STATE Num:65 Check Scan Retry Count Over Or Not
   RUNG wire#powerrail
      Contact( #s65_ChkScanRetryOver )
      wire#w1
      I_Contact( #s65_ChkScanRetryOver_T1 )
      I_Contact( #s65_ChkScanRetryOver_T2 )
      wire#w2
      Coil( #s65_ChkScanRetryOver )
   END_RUNG
   RUNG wire#powerrail
      Contact( #s52_WaitScanOver_T2 )
   END_RUNG wire#w1
   RUNG wire#w2
      { S7_GenerateENO := "TRUE" } Move(in := 65, out1 => #StateNo)
   END_RUNG
   // the same network as SCL:
   #s65_ChkScanRetryOver := (#s65_ChkScanRetryOver OR #s52_WaitScanOver_T2) AND NOT #s65_ChkScanRetryOver_T1 AND NOT #s65_ChkScanRetryOver_T2;
   IF #s65_ChkScanRetryOver THEN #StateNo := 65; END_IF;
END_REGION

NETWORK
TITLE = Actions for STATE Num:65 Check Scan Retry Count Over Or Not
      A     #s65_ChkScanRetryOver_T1;
      L     #sScanRetryCount;
      L     1;
      +I;
      T     #sScanRetryCount;

REGION Network 55: Transition for STATE Num:66 Wait for Operator desicion
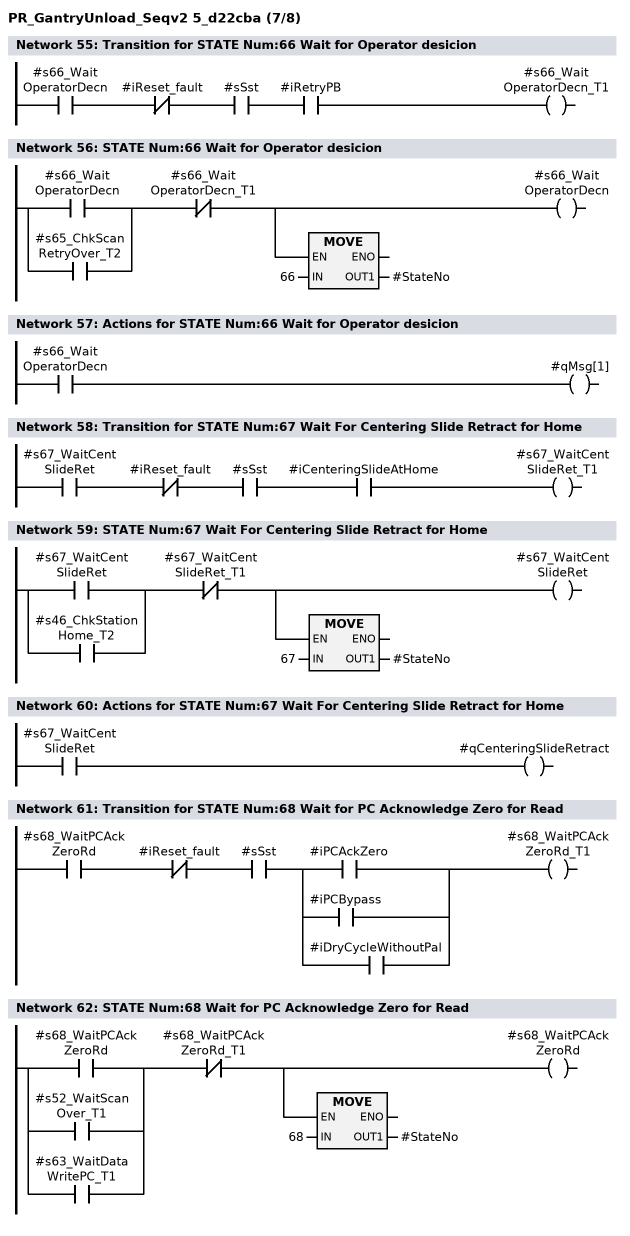
   RUNG wire#powerrail
      Contact( #s66_WaitOperatorDecn )
      I_Contact( #iReset_fault )
      Contact( #sSst )
      Contact( #iRetryPB )
      Coil( #s66_WaitOperatorDecn_T1 )
   END_RUNG
   // the same network as SCL:
   #s66_WaitOperatorDecn_T1 := #s66_WaitOperatorDecn AND NOT #iReset_fault AND #sSst AND #iRetryPB;
END_REGION

REGION Network 56: STATE Num:66 Wait for Operator desicion
   RUNG wire#powerrail
      Contact( #s66_WaitOperatorDecn )
      wire#w1
      I_Contact( #s66_WaitOperatorDecn_T1 )
      wire#w2
      Coil( #s66_WaitOperatorDecn )
   END_RUNG
   RUNG wire#powerrail
      Contact( #s65_ChkScanRetryOver_T2 )
   END_RUNG wire#w1
   RUNG wire#w2
      { S7_GenerateENO := "TRUE" } Move(in := 66, out1 => #StateNo)
   END_RUNG
   // the same network as SCL:
   #s66_WaitOperatorDecn := (#s66_WaitOperatorDecn OR #s65_ChkScanRetryOver_T2) AND NOT #s66_WaitOperatorDecn_T1;
   IF #s66_WaitOperatorDecn THEN #StateNo := 66; END_IF;
END_REGION

REGION Network 57: Actions for STATE Num:66 Wait for Operator desicion
   RUNG wire#powerrail
      Contact( #s66_WaitOperatorDecn )
      Coil( #qMsg[1] )
   END_RUNG
   // the same network as SCL:
   #qMsg[1] := #s66_WaitOperatorDecn;
END_REGION

REGION Network 58: Transition for STATE Num:67 Wait For Centering Slide Retract for Home
   RUNG wire#powerrail
      Contact( #s67_WaitCentSlideRet )
      I_Contact( #iReset_fault )
      Contact( #sSst )
      Contact( #iCenteringSlideAtHome )
      Coil( #s67_WaitCentSlideRet_T1 )
   END_RUNG
   // the same network as SCL:
   #s67_WaitCentSlideRet_T1 := #s67_WaitCentSlideRet AND NOT #iReset_fault AND #sSst AND #iCenteringSlideAtHome;
END_REGION

REGION Network 59: STATE Num:67 Wait For Centering Slide Retract for Home
   RUNG wire#powerrail
      Contact( #s67_WaitCentSlideRet )
      wire#w1
      I_Contact( #s67_WaitCentSlideRet_T1 )
      wire#w2
      Coil( #s67_WaitCentSlideRet )
   END_RUNG
   RUNG wire#powerrail
      Contact( #s46_ChkStationHome_T2 )
   END_RUNG wire#w1
   RUNG wire#w2
      { S7_GenerateENO := "TRUE" } Move(in := 67, out1 => #StateNo)
   END_RUNG
   // the same network as SCL:
   #s67_WaitCentSlideRet := (#s67_WaitCentSlideRet OR #s46_ChkStationHome_T2) AND NOT #s67_WaitCentSlideRet_T1;
   IF #s67_WaitCentSlideRet THEN #StateNo := 67; END_IF;
END_REGION

REGION Network 60: Actions for STATE Num:67 Wait For Centering Slide Retract for Home
   RUNG wire#powerrail
      Contact( #s67_WaitCentSlideRet )
      Coil( #qCenteringSlideRetract )
   END_RUNG
   // the same network as SCL:
   #qCenteringSlideRetract := #s67_WaitCentSlideRet;
END_REGION

REGION Network 61: Transition for STATE Num:68 Wait for PC Acknowledge Zero for Read
   RUNG wire#powerrail
      Contact( #s68_WaitPCAckZeroRd )
      I_Contact( #iReset_fault )
      Contact( #sSst )
      wire#w1
      Contact( #iPCAckZero )
      wire#w2
      Coil( #s68_WaitPCAckZeroRd_T1 )
   END_RUNG
   RUNG wire#w1
      Contact( #iPCBypass )
   END_RUNG wire#w2
   RUNG wire#w1
      Contact( #iDryCycleWithoutPal )
   END_RUNG wire#w2
   // the same network as SCL:
   #s68_WaitPCAckZeroRd_T1 := #s68_WaitPCAckZeroRd AND NOT #iReset_fault AND #sSst AND (#iPCAckZero OR #iPCBypass OR #iDryCycleWithoutPal);
END_REGION

REGION Network 62: STATE Num:68 Wait for PC Acknowledge Zero for Read
   RUNG wire#powerrail
      Contact( #s68_WaitPCAckZeroRd )
      wire#w1
      I_Contact( #s68_WaitPCAckZeroRd_T1 )
      wire#w2
      Coil( #s68_WaitPCAckZeroRd )
   END_RUNG
   RUNG wire#powerrail
      Contact( #s52_WaitScanOver_T1 )
   END_RUNG wire#w1
   RUNG wire#powerrail
      Contact( #s63_WaitDataWritePC_T1 )
   END_RUNG wire#w1
   RUNG wire#w2
      { S7_GenerateENO := "TRUE" } Move(in := 68, out1 => #StateNo)
   END_RUNG
   // the same network as SCL:
   #s68_WaitPCAckZeroRd := (#s68_WaitPCAckZeroRd OR #s52_WaitScanOver_T1 OR #s63_WaitDataWritePC_T1) AND NOT #s68_WaitPCAckZeroRd_T1;
   IF #s68_WaitPCAckZeroRd THEN #StateNo := 68; END_IF;
END_REGION

REGION Network 63: Transition for STATE Num:69 Wait for Data Read Over From PC
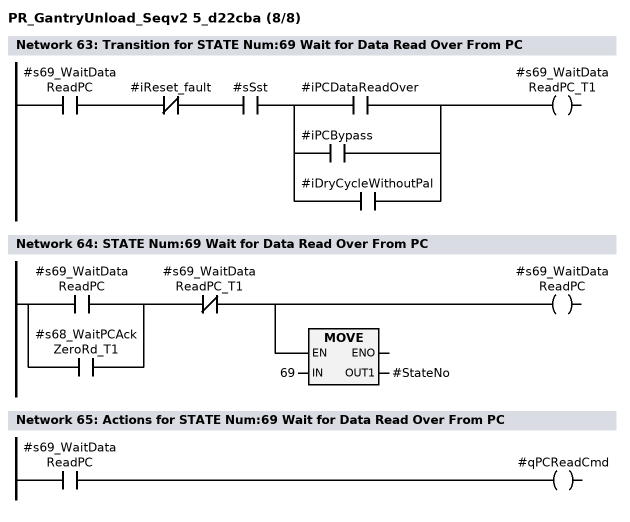
   RUNG wire#powerrail
      Contact( #s69_WaitDataReadPC )
      I_Contact( #iReset_fault )
      Contact( #sSst )
      wire#w1
      Contact( #iPCDataReadOver )
      wire#w2
      Coil( #s69_WaitDataReadPC_T1 )
   END_RUNG
   RUNG wire#w1
      Contact( #iPCBypass )
   END_RUNG wire#w2
   RUNG wire#w1
      Contact( #iDryCycleWithoutPal )
   END_RUNG wire#w2
   // the same network as SCL:
   #s69_WaitDataReadPC_T1 := #s69_WaitDataReadPC AND NOT #iReset_fault AND #sSst AND (#iPCDataReadOver OR #iPCBypass OR #iDryCycleWithoutPal);
END_REGION

REGION Network 64: STATE Num:69 Wait for Data Read Over From PC
   RUNG wire#powerrail
      Contact( #s69_WaitDataReadPC )
      wire#w1
      I_Contact( #s69_WaitDataReadPC_T1 )
      wire#w2
      Coil( #s69_WaitDataReadPC )
   END_RUNG
   RUNG wire#powerrail
      Contact( #s68_WaitPCAckZeroRd_T1 )
   END_RUNG wire#w1
   RUNG wire#w2
      { S7_GenerateENO := "TRUE" } Move(in := 69, out1 => #StateNo)
   END_RUNG
   // the same network as SCL:
   #s69_WaitDataReadPC := (#s69_WaitDataReadPC OR #s68_WaitPCAckZeroRd_T1) AND NOT #s69_WaitDataReadPC_T1;
   IF #s69_WaitDataReadPC THEN #StateNo := 69; END_IF;
END_REGION

REGION Network 65: Actions for STATE Num:69 Wait for Data Read Over From PC
   RUNG wire#powerrail
      Contact( #s69_WaitDataReadPC )
      Coil( #qPCReadCmd )
   END_RUNG
   // the same network as SCL:
   #qPCReadCmd := #s69_WaitDataReadPC;
END_REGION
END_FUNCTION_BLOCK
